(* IEC 61131-3 sources: Elmo_Master/Lasal_PRG/Elmo_EtherCAT_Test_4Axis/Network/Comm_Network, 1 file *)

(* ---- ONE_Comm_Network_Table.st ---- *)
#define OBJECTS_CONFIG

//Define part of class _TCPIPServer
#ifndef OS_VERSION_MIN_SALAMANDER
    #define OS_VERSION_MIN_SALAMANDER          0x9000
  #endif
  #define TCP_SVR_NO_ERROR                          0

  #define TCP_SVR_ERR_INVALID_SOCKET            -1

  #define TCP_SVR_ERR_SET_PARA_INVALID_CMD     -10
  #define TCP_SVR_ERR_SET_PARA_INVALID_SUB_CMD -11

  #define TCP_SVR_ERR_TASK_ALREADY_EXIST       -12

  // - RETURN VALUES PRIVATE METHOD Read_AP_TaskPeriod
  #define TCP_SVR_ERR_TASK_TIME_NO_APP            -31
  #define TCP_SVR_ERR_TASK_TIME_WRONG_TASK_TYPE   -33
  #define TCP_SVR_ERR_TASK_TIME_OBJ_NOT_FOUND     -35

  // - RETURN VALUES PRIVATE METHOD Read_LSLOBJ_CRC32
  #define TCP_SVR_ERR_GET_LSLOBJ_NAME             -20
  #define TCP_SVR_ERR_INVALID_POINTER             -21

  // - RETURN VALUES PRIVATE METHOD AP_TaskCreate
  #define TCP_SVR_ERR_TASK_CREATE                 -40

  // - RETURN VALUES PRIVATE METHOD AP_SemaCreate
  #define TCP_SVR_ERR_SEMA_CREATE                 -50
  #define TCP_SVR_ERR_SEMA_INVALID_IDX            -51
  #define TCP_SVR_ERR_SEMA_INVALID_NAME           -52

  #define TCP_SVR_SEND_BUFFER_EMPTY               -6
  #define TCP_SVR_ERR_SEND_BUFFER_FATAL_ERROR     -7

  #define TCP_SVR_SEND_BUFFER_FULL      -4

  #define TCP_SVR_SOCK_INFO_CONNECT                 1
  #define TCP_SVR_SOCK_INFO_DISCONNECT              0

  #define TCP_SVR_ERR_GROUP_OS                      0
  #define TCP_SVR_ERR_GROUP_AP                      1

  #define TCP_SVR_ERR_CODE_AP_TIMEOUT              -1

  #ifndef INIT_FIRSTSCAN
    #define INIT_FIRSTSCAN                         12
  #endif

  #ifndef AP_TASK_PRIORITY_DEFAULT
    #define AP_TASK_PRIORITY_DEFAULT               14
  #endif

  #define TCP_SVR_ERR_MAIN_INIT                   -90

  #define TCP_SVR_ERR_MAX_CONN                    -80

  #ifndef KEEPALIVE_INTERVAL_DEFAULT
    #define KEEPALIVE_INTERVAL_DEFAULT           7200
  #endif

  #ifndef KEEPALIVE_RETRYTIME_DEFAULT
    #define KEEPALIVE_RETRYTIME_DEFAULT            75
  #endif

  #ifndef KEEPALIVE_RETRYCNT_DEFUALT
    #define KEEPALIVE_RETRYCNT_DEFUALT             10
  #endif

  #ifndef CLOSE_SOCKET_TYPE_DEFAULT
    #define CLOSE_SOCKET_TYPE_DEFAULT               0
  #endif
#include "..\..\Class\_TCPIPServer\_TCPIPServer.h"
#include "..\..\Class\_TCPIPServer\SalamanderDelay.h"
//Define part of class _UDPTransceiver
#define UDP_MAX_SOCKETS               6                             // Max number of socket

#define UDP_CLT_SEND_OK               0                             // Send ok
#define UDP_CLT_INVALID_HANDLE        -1                            // Invalid handle
#define UDP_CLT_NOT_OPEN              -2                            // Socket is not open
#define UDP_CLT_SEND_FAILED           -3                            // Send failed
#define UDP_CLT_SEND_BUFFER_FULL      -4                            // Send buffer is full
#define UDP_CLT_DATA_TO_BIG           -5                            // Data to big
#define UDP_CLT_INVALID_DATA          -6

#define UDP_MAXIMUM_SEGMENT_SIZE      1452                          //

#define MAX_MSG_CYC_SEND                5
#define MAX_MSG_CYC_RECV                5

#define UDP_CLT_INFO_ADDED          0
#define UDP_CLT_INFO_BOUND          1
#define UDP_CLT_INFO_CLOSED         2
//Define part of class LMCUdpCallbackSender
#ifndef LMC_UDP_CALLBACK_ENABLE_LEGACY_FIXTURE
#define LMC_UDP_CALLBACK_ENABLE_LEGACY_FIXTURE 0
#endif
#include <.\lsl_st_mt.h>

FUNCTION GLOBAL TAB ONE_Comm_Network
-1$UINT, 0$UINT,
0$UINT, 0$UINT,

16$UDINT,
TO_UDINT(916194998), "_CheckSum", 1$UINT, 0$UINT, 2$UINT,
TO_UDINT(4107457475), "_TCPIPServer", 1$UINT, 2$UINT, 0$UINT,
TO_UDINT(3417437475), "_TCPIPServerInterface", 1$UINT, 1$UINT, 0$UINT,
TO_UDINT(3808005437), "_UDPTransceiver", 1$UINT, 2$UINT, 1$UINT,
TO_UDINT(3441197119), "_UDPTransceiverInterface", 1$UINT, 3$UINT, 0$UINT,
TO_UDINT(794617671), "CriticalSection", 0$UINT, 4$UINT, 2$UINT,
TO_UDINT(4292381624), "LMCControlCommandService", 0$UINT, 0$UINT, 1$UINT,
TO_UDINT(1037074496), "LMCDiagnosticsService", 0$UINT, 0$UINT, 1$UINT,
TO_UDINT(2393574248), "LMCSetPositionStore", 0$UINT, 0$UINT, 1$UINT,
TO_UDINT(287734476), "LMCUdpCallbackSender", 0$UINT, 0$UINT, 1$UINT,
TO_UDINT(2225119864), "MerkerEx", 1$UINT, 22$UINT, 3$UINT,
TO_UDINT(1850111279), "String", 1$UINT, 11$UINT, 3$UINT,
TO_UDINT(2898603620), "StringInternal", 1$UINT, 86$UINT, 0$UINT,
TO_UDINT(2859426109), "TCPIPServer", 0$UINT, 0$UINT, 1$UINT,
TO_UDINT(684024945), "TCPMotionInterface", 0$UINT, 0$UINT, 1$UINT,
TO_UDINT(3232495061), "VirtualBaseInit", 1$UINT, 3$UINT, 0$UINT,

_NO_ATTR, TO_UDINT(1739067253), "LMCSETPOSITIONCHECKSUM1",
1$UINT, TO_UDINT(4285366611), "TCPIPSERVER1\_BASE\CHECKSUM",

_NO_ATTR, TO_UDINT(4169137385), "LMCUDPTRANSCEIVER1",

1$UINT, TO_UDINT(857947721), "LMCUDPCALLBACKSENDER1\_BASE\CRITICALSECTION_UDP",
1$UINT, TO_UDINT(1512526909), "LMCUDPTRANSCEIVER1\CRITICALSECTION_UDP",

_NO_ATTR, TO_UDINT(1184435330), "LMCCONTROLCOMMANDSERVICE1",

_NO_ATTR, TO_UDINT(4114448039), "LMCDIAGNOSTICSSERVICE1",

_NO_ATTR, TO_UDINT(3225136598), "LMCSETPOSITIONSTORE1",

_NO_ATTR, TO_UDINT(287262550), "LMCUDPCALLBACKSENDER1",

1$UINT, TO_UDINT(2143358748), "TCPIPSERVER1\_BASE\STRSEMANAME01\MERKEREX0",
1$UINT, TO_UDINT(3861080349), "TCPIPSERVER1\_BASE\STRSEMANAME02\MERKEREX0",
1$UINT, TO_UDINT(3045102150), "TCPIPSERVER1\_BASE\STRTASKNAME\MERKEREX0",

1$UINT, TO_UDINT(1660672605), "TCPIPSERVER1\_BASE\STRSEMANAME01",
1$UINT, TO_UDINT(4226976743), "TCPIPSERVER1\_BASE\STRSEMANAME02",
1$UINT, TO_UDINT(4139250991), "TCPIPSERVER1\_BASE\STRTASKNAME",

_NO_ATTR, TO_UDINT(3676228807), "TCPIPSERVER1",

_NO_ATTR, TO_UDINT(2767612793), "TCPMOTIONINTERFACE1",

//Internal connections
0$UDINT,
9$UDINT,
TO_UDINT(2), "CriticalSection_UDP", TO_UDINT(4),
TO_UDINT(8), "CriticalSection_UDP", TO_UDINT(3),
TO_UDINT(12), "MerkerEx0", TO_UDINT(9),
TO_UDINT(13), "MerkerEx0", TO_UDINT(10),
TO_UDINT(14), "MerkerEx0", TO_UDINT(11),
TO_UDINT(15), "CheckSum", TO_UDINT(1),
TO_UDINT(15), "StrTaskName", TO_UDINT(14),
TO_UDINT(15), "StrSemaName01", TO_UDINT(12),
TO_UDINT(15), "StrSemaName02", TO_UDINT(13),
0$UDINT,
11$UDINT,
TO_UDINT(5), "SetPositionStore", TO_UDINT(7), "ClassSvr",
TO_UDINT(6), "AxisOwnership", TO_UDINT(5), "ClassSvr",
TO_UDINT(7), "CheckSum", TO_UDINT(0), "ClassSvr",
TO_UDINT(8), "_UDPTransceiver", TO_UDINT(2), "sControl",
TO_UDINT(12), "DataBuffer", TO_UDINT(9), "m_udLength",
TO_UDINT(13), "DataBuffer", TO_UDINT(10), "m_udLength",
TO_UDINT(14), "DataBuffer", TO_UDINT(11), "m_udLength",
TO_UDINT(16), "_TCPIPServer", TO_UDINT(15), "Control",
TO_UDINT(16), "Diagnostics", TO_UDINT(6), "ClassSvr",
TO_UDINT(16), "ControlCommands", TO_UDINT(5), "ClassSvr",
TO_UDINT(16), "CallbackSender", TO_UDINT(8), "ClassSvr",

//Initialization values
0$UDINT,
23$UDINT,
TO_UDINT(2), "cSizeOfTXBuffer", TO_UDINT(8 kb),//|Comm_Network.LMCUdpTransceiver1.cSizeOfTXBuffer;
TO_UDINT(2), "cSizeOfRXBuffer", TO_UDINT(512),//|Comm_Network.LMCUdpTransceiver1.cSizeOfRXBuffer;
TO_UDINT(5), "AxisRebaseRequiredState", TO_UDINT(16#5242530F),//|Comm_Network.LMCControlCommandService1.AxisRebaseRequiredState;
TO_UDINT(6), "DiagnosticsBootCounter", TO_UDINT(0),//|Comm_Network.LMCDiagnosticsService1.DiagnosticsBootCounter;
TO_UDINT(8), "QueueDepth", TO_UDINT(0),//|Comm_Network.LMCUdpCallbackSender1.QueueDepth;
TO_UDINT(8), "QueuedCount", TO_UDINT(0),//|Comm_Network.LMCUdpCallbackSender1.QueuedCount;
TO_UDINT(8), "RingAcceptedCount", TO_UDINT(0),//|Comm_Network.LMCUdpCallbackSender1.RingAcceptedCount;
TO_UDINT(8), "AdmissionRetryCount", TO_UDINT(0),//|Comm_Network.LMCUdpCallbackSender1.AdmissionRetryCount;
TO_UDINT(8), "QueueFullDropCount", TO_UDINT(0),//|Comm_Network.LMCUdpCallbackSender1.QueueFullDropCount;
TO_UDINT(8), "AdmissionErrorDropCount", TO_UDINT(0),//|Comm_Network.LMCUdpCallbackSender1.AdmissionErrorDropCount;
TO_UDINT(8), "DisarmClearedCount", TO_UDINT(0),//|Comm_Network.LMCUdpCallbackSender1.DisarmClearedCount;
TO_UDINT(8), "TransportErrorCount", TO_UDINT(0),//|Comm_Network.LMCUdpCallbackSender1.TransportErrorCount;
TO_UDINT(8), "LastAdmissionResult", TO_UDINT(0),//|Comm_Network.LMCUdpCallbackSender1.LastAdmissionResult;
TO_UDINT(9), "ThreadSafe", TO_UDINT(0),//|Comm_Network.StrSemaName01\_base\TCPIPServer1\MerkerEx0.ThreadSafe;
TO_UDINT(10), "ThreadSafe", TO_UDINT(0),//|Comm_Network.StrSemaName02\_base\TCPIPServer1\MerkerEx0.ThreadSafe;
TO_UDINT(11), "ThreadSafe", TO_UDINT(0),//|Comm_Network.StrTaskName\_base\TCPIPServer1\MerkerEx0.ThreadSafe;
TO_UDINT(12), "SingleRealloc", TO_UDINT(1),//|Comm_Network._base\TCPIPServer1\StrSemaName01.SingleRealloc;
TO_UDINT(13), "SingleRealloc", TO_UDINT(1),//|Comm_Network._base\TCPIPServer1\StrSemaName02.SingleRealloc;
TO_UDINT(14), "SingleRealloc", TO_UDINT(1),//|Comm_Network._base\TCPIPServer1\StrTaskName.SingleRealloc;
TO_UDINT(15), "Port", TO_UDINT(4000),//|Comm_Network.TCPIPServer1.Port;
TO_UDINT(15), "MaxConnections", TO_UDINT(2),//|Comm_Network.TCPIPServer1.MaxConnections;
TO_UDINT(15), "ConnectionsPerRun", TO_UDINT(1),//|Comm_Network.TCPIPServer1.ConnectionsPerRun;
TO_UDINT(15), "Config", TO_UDINT(0),//|Comm_Network.TCPIPServer1.Config;

//Symbolic initialization values
0$UDINT,
0$UDINT,

//Initialization of string values
0$UDINT,
0$UDINT,

//Configuration of tasks (RealTime, Cyclic, Background)
0$UDINT,
0$UDINT,

0$UDINT,
4$UDINT,
TO_UDINT(2), (10)$UDINT, 4194303$DINT, 	//LMCUDPTRANSCEIVER1
TO_UDINT(8), (10)$UDINT, 4194303$DINT, 	//LMCUDPCALLBACKSENDER1
TO_UDINT(15), (1)$UDINT, 4194303$DINT, 	//TCPIPSERVER1
TO_UDINT(16), (1)$UDINT, 4194303$DINT, 	//TCPMOTIONINTERFACE1

0$UDINT,
0$UDINT,

//External connections
0$UDINT,
17$UDINT,
TO_UDINT(5), "InputLatch", C_DIR, TO_UDINT(3311388916), "LMCEcatInputLatch1","ClassSvr",
TO_UDINT(5), "LMCAxis1", C_DIR, TO_UDINT(1307168646), "_LMCAxis1","Control",
TO_UDINT(5), "LMCAxis2", C_DIR, TO_UDINT(3571490364), "_LMCAxis2","Control",
TO_UDINT(5), "LMCAxis3", C_DIR, TO_UDINT(2749869738), "_LMCAxis3","Control",
TO_UDINT(5), "LMCAxis4", C_DIR, TO_UDINT(1032010505), "_LMCAxis4","Control",
TO_UDINT(5), "LMCAxis5", C_DIR, TO_UDINT(1250167711), "_LMCAxis5","Control",
TO_UDINT(5), "LMCAxis6", C_DIR, TO_UDINT(3549256229), "_LMCAxis6","Control",
TO_UDINT(5), "LMCAxis7", C_DIR, TO_UDINT(2760534707), "_LMCAxis7","Control",
TO_UDINT(5), "LMCAxis8", C_DIR, TO_UDINT(875919138), "_LMCAxis8","Control",
TO_UDINT(5), "LMCAxis9", C_DIR, TO_UDINT(1127368628), "_LMCAxis9","Control",
TO_UDINT(5), "LMCRobot", C_DIR, TO_UDINT(669706412), "_LMCRobotBase1","Control",
TO_UDINT(6), "InputLatch", C_DIR, TO_UDINT(3311388916), "LMCEcatInputLatch1","ClassSvr",
TO_UDINT(6), "RecorderStore", C_DIR, TO_UDINT(1161287402), "LMCRecorderStore1","ClassSvr",
TO_UDINT(6), "SdoAxis1", C_DIR, TO_UDINT(1999418485), "LMCSdoExecutor1","ClassState",
TO_UDINT(6), "SdoAxis2", C_DIR, TO_UDINT(3995461071), "LMCSdoExecutor2","ClassState",
TO_UDINT(6), "SdoAxis3", C_DIR, TO_UDINT(2569196889), "LMCSdoExecutor3","ClassState",
TO_UDINT(6), "SdoAxis4", C_DIR, TO_UDINT(122044666), "LMCSdoExecutor4","ClassState",

//Magic internal connections
0$UDINT,
0$UDINT,

//Configuration of timeslots of tasks (RealTime, Cyclic)
#ifdef __LSLLDR_TIMESLOTS__
0$UDINT,
0$UDINT,

0$UDINT,
0$UDINT,

#endif //__LSLLDR_TIMESLOTS__

//MultiMaster connections
#ifdef __LSLLDR_MULTIMASTER__
0$UDINT,
0$UDINT,
#endif //__LSLLDR_MULTIMASTER__

//Configuration for task ID (RealTime, CyclicTime)
#ifdef __LSLLDR_TASKID__
"\\\\TASKS2  "
0$UDINT,
0$UDINT,

0$UDINT,
4$UDINT,
(0)$UDINT, 	//LMCUDPTRANSCEIVER1
(0)$UDINT, 	//LMCUDPCALLBACKSENDER1
(0)$UDINT, 	//TCPIPSERVER1
(0)$UDINT, 	//TCPMOTIONINTERFACE1

0$UDINT,
0$UDINT,

#endif //__LSLLDR_TASKID__

END_FUNCTION
